(* IEC 61131-3 sources: test/Class/AI040 (part 2) *)

    //if raw values is selected dont correct gain factor
    if sScaleSettings.bRawValue.Channel4 = TRUE then
      dTempGain := 1;
    end_if;

    sWriteCalibData.Divisor.Channel4    := sReadCalibData.Channel4[dTempArray].Divisor;
    sWriteCalibData.Multiplier.Channel4 := sReadCalibData.Channel4[dTempArray].Multiplier;
    sWriteCalibData.Offset.Channel4     := sReadCalibData.Channel4[dTempArray].Offset;
    //if there is no valid calib data set it to mul and div to 1
    if sWriteCalibData.Divisor.Channel4 = 0 then
      sWriteCalibData.Divisor.Channel4    := 1;
      sWriteCalibData.Multiplier.Channel4 := 1;
      sWriteCalibData.Offset.Channel4     := 0;
    end_if;
  end_if;

END_FUNCTION

FUNCTION VIRTUAL GLOBAL AI040::DisconnectEvent

  SdiasBase::DisconnectEvent();

END_FUNCTION

FUNCTION AI040::SetScale
VAR_OUTPUT
  eModuleInitState 	: iprStates;
END_VAR
VAR
	dScale : DINT;
END_VAR

  eModuleInitState := READY;

  //analog input 1
  //*************************************************************************************************************
  if sMeasureControl.ArrayAssignment.ChArrayActivated.Channel1 then
    AI1MaxValue  := AI1MaxValue.Read();
    AI1MinValue  := AI1MinValue.Read();

    //check if calculation is necessary
    if ((AI1MaxValue <> AI040_FIRMWARE_MAX) | (AI1MinValue <> AI040_FIRMWARE_MIN)) then

      ScaleAI1 := TRUE;

      dScale := AI1MaxValue-AI1MinValue;

      if dScale = 0 then
        eModuleInitState := ERROR;
        eInitState := _InvalidConfguration;
        LogValue("@014C (AI040::SetScale) Invalid minimal and maximal value settings for channel {0}. The values must not be the same.",1);
        return;
      end_if;

      sScaleSettings.Multiplier.Channel1 := dScale;
      sScaleSettings.Divider.Channel1 := (AI040_FIRMWARE_MAX - AI040_FIRMWARE_MIN);
      sScaleSettings.Offset.Channel1  := (AI1MinValue * sScaleSettings.Divider.Channel1)/(sScaleSettings.Multiplier.Channel1) - AI040_FIRMWARE_MIN;
    else
      sScaleSettings.Offset.Channel1 := 0;
    end_if;
  end_if;

  //analog input 2
  //*************************************************************************************************************
  if sMeasureControl.ArrayAssignment.ChArrayActivated.Channel2 then
    AI2MaxValue  := AI2MaxValue.Read();
    AI2MinValue  := AI2MinValue.Read();

    //check if calculation is necessary
    if ((AI2MaxValue <> AI040_FIRMWARE_MAX) | (AI2MinValue <> AI040_FIRMWARE_MIN)) then

      ScaleAI2 := TRUE;

      dScale := AI2MaxValue-AI2MinValue;

      if dScale = 0 then
        eModuleInitState := ERROR;
        eInitState := _InvalidConfguration;
        LogValue("@014C (AI040::SetScale) Invalid minimal and maximal value settings for channel {0}. The values must not be the same.",2);
        return;
      end_if;

      sScaleSettings.Multiplier.Channel2 := dScale;
      sScaleSettings.Divider.Channel2 := (AI040_FIRMWARE_MAX - AI040_FIRMWARE_MIN);
      sScaleSettings.Offset.Channel2  := (AI2MinValue * sScaleSettings.Divider.Channel2)/(sScaleSettings.Multiplier.Channel2) - AI040_FIRMWARE_MIN;
    else
      sScaleSettings.Offset.Channel2 := 0;
    end_if;
  end_if;

  //analog input 3
  //*************************************************************************************************************
  if sMeasureControl.ArrayAssignment.ChArrayActivated.Channel3 then
    AI3MaxValue  := AI3MaxValue.Read();
    AI3MinValue  := AI3MinValue.Read();

    //check if calculation is necessary
    if ((AI3MaxValue <> AI040_FIRMWARE_MAX) | (AI3MinValue <> AI040_FIRMWARE_MIN)) then

      ScaleAI3 := TRUE;

      dScale := AI3MaxValue-AI3MinValue;

      if dScale = 0 then
        eModuleInitState := ERROR;
        eInitState := _InvalidConfguration;
        LogValue("@014C (AI040::SetScale) Invalid minimal and maximal value settings for channel {0}. The values must not be the same.",3);
        return;
      end_if;

      sScaleSettings.Multiplier.Channel3 := dScale;
      sScaleSettings.Divider.Channel3    := (AI040_FIRMWARE_MAX - AI040_FIRMWARE_MIN);
      sScaleSettings.Offset.Channel3     := (AI3MinValue * sScaleSettings.Divider.Channel3)/(sScaleSettings.Multiplier.Channel3) - AI040_FIRMWARE_MIN;
    else
      sScaleSettings.Offset.Channel3 := 0;
    end_if;
  end_if;

  //analog input 4
  //*************************************************************************************************************
  if sMeasureControl.ArrayAssignment.ChArrayActivated.Channel4 then
    AI4MaxValue  := AI4MaxValue.Read();
    AI4MinValue  := AI4MinValue.Read();

    //check if calculation is necessary
    if ((AI4MaxValue <> AI040_FIRMWARE_MAX) | (AI4MinValue <> AI040_FIRMWARE_MIN)) then

      ScaleAI4 := TRUE;

      dScale := AI4MaxValue-AI4MinValue;

      if dScale = 0 then
        eModuleInitState := ERROR;
        eInitState := _InvalidConfguration;
        LogValue("@014C (AI040::SetScale) Invalid minimal and maximal value settings for channel {0}. The values must not be the same.",4);
        return;
      end_if;

      sScaleSettings.Multiplier.Channel4 := dScale;
      sScaleSettings.Divider.Channel4    := (AI040_FIRMWARE_MAX - AI040_FIRMWARE_MIN);
      sScaleSettings.Offset.Channel4     := (AI4MinValue * sScaleSettings.Divider.Channel4)/(sScaleSettings.Multiplier.Channel4) - AI040_FIRMWARE_MIN;
    else
      sScaleSettings.Offset.Channel4 := 0;
    end_if;
  end_if;

END_FUNCTION

FUNCTION VIRTUAL GLOBAL AI040::ClassState::NewInst
	VAR_INPUT
		pPara 	: ^CmdStruct;
		pResult 	: ^Results;
	END_VAR
	VAR_OUTPUT
		ret_code 	: IprStates;
	END_VAR
  VAR
  	udActDataCount  : UDINT;
  END_VAR

	CASE pPara^.uiCmd OF
//**********************************************************************************************************************************************************
    SDIAS_CLT_GET_ANALOG_DATA_BUFFER:
      // init with error, ok is set later
      ret_code := ERROR;

      if pPara^.aPara[0] = 1 then
        // request is version 1

        // check valid channel nr
        if (pPara^.aPara[1] >= 1) & (pPara^.aPara[1] <= 4) then

          // init result
          ret_code := READY;
          pResult^.aData[0x0]       := 1; //version 1
          pResult^.aData[0x1]       := AI040_SIZE_ONE_VALUE;
          pResult^.aData[0x2]$UDINT := to_udint(uiMaxValuesCycle);
          pResult^.aData[0x6]$UDINT := 0; // copied amount is set later
          pResult^.aData[0xA]$UDINT := 0; // no counter
          pResult^.aData[0xB]$UDINT := 0; // so set counter to 0

          // copy requested data amount, limit to avaliable data
          if (pPara^.aPara[2] <> NIL) & (pPara^.aPara[3]$UDINT > 0) then
            udActDataCount := pPara^.aPara[3]$UDINT;
            if (udActDataCount AND 1) = 1 then
              udActDataCount -= 1; // only whole values
            end_if;
            if udActDataCount > (uiMaxValuesCycle*AI040_SIZE_ONE_VALUE) then
              udActDataCount := (uiMaxValuesCycle*AI040_SIZE_ONE_VALUE);
            end_if;
            if GetData(usChannelNr:= pPara^.aPara[1]$USINT, uiDataLength:=udActDataCount$UINT, pBufferData:=pPara^.aPara[2]$^INT) = 0 then
              pResult^.aData[6]$UDINT := udActDataCount / AI040_SIZE_ONE_VALUE;
            //else
              // no data copied, probably data is INVALID
            end_if;
          //else
            //no data requested
          end_if;
        //else
          // wrong channel
        end_if;
      //else
        // unknown version of the request
      end_if;

//**********************************************************************************************************************************************************
  ELSE
    // we forward this message to the base class
		ret_code := SdiasBase::NewInst(pPara, pResult);
	END_CASE;

END_FUNCTION
